Staubli VAL3: utBorder.dtx

public string sBorderColour
public string sBorderStyle
public string sBorderWidth
